FUNCTION "LGF_MatrixInverse" : Void
{ S7_Optimized_Access := 'TRUE' }
AUTHOR : Siemens_Digital_Industry
FAMILY : LGF
NAME : LGF_MatrixInverse
   VAR_OUTPUT
      error : Bool;
      status : Word;
   END_VAR

   VAR_IN_OUT
      matrix : Array[*, *] of LReal;
      matrixResult : Array[*, *] of LReal;
   END_VAR

   VAR_TEMP
      tempMatrix1LowerBoundRows : DInt;
      tempMatrix1LowerBoundColumns : DInt;
      tempMatrix1UpperBoundRows : DInt;
      tempMatrix1UpperBoundColumns : DInt;
      tempResultMatrixLowerBoundRows : DInt;
      tempResultMatrixLowerBoundColumns : DInt;
      tempResultMatrixUpperBoundRows : DInt;
      tempResultMatrixUpperBoundColumns : DInt;
      tempCounterRows : DInt;
      tempCounterColumns : DInt;
      tempColumns : DInt;
      tempRows : DInt;
      tempK : DInt;
      tempI : DInt;
      tempJ : DInt;
      tempMatrixElement : LReal;
   END_VAR

   VAR CONSTANT
      PRECISION : LReal := 1.0E-10;
      NEGATIVE_NUMERATOR : LReal := -1.0;
      ZERO : UInt := 0;
      ONE : UInt := 1;
      ROWS : UInt := 1;
      COLUMNS : UInt := 2;
      STATUS_NO_ERROR : Word := 16#0000;
      ERR_NOT_SQUARE_MATRIX : Word := 16#8200;
      ERR_ALGORITHM_NOT_POSSIBLE : Word := 16#8201;
      ERR_MATR1_LOWBOUND_ROWS_RESMATR_LOWBOUND_ROWS : Word := 16#8202;
      ERR_MATR1_LOWBOUND_COLUMNS_RESMATR_LOWBOUND_COLUMNS : Word := 16#8203;
      ERR_MATR1_UPPBOUND_ROWS_RESMATR_UPPBOUND_ROWS : Word := 16#8204;
      ERR_MATR1_UPPBOUND_COLUMNS_RESMATR_UPPBOUND_COLUMNS : Word := 16#8205;
   END_VAR


BEGIN
	REGION Block info header
	  //=============================================================================
	  // SIEMENS AG / (c)Copyright 2017
	  //-------------------------------------------------------------------------------
	  // Title:            LGF_MatrixInverse
	  // Comment/Function: Caluclates an inverted version of a matrix
	  // Library/Family:   LGF(Library General Functions)
	  // Author:           Siemens Digital Industry Support
	  // Tested with:      S7-PLCSIM Advanced V2.0 SP1
	  // Engineering:      TIA Portal V15 Update 2
	  // Restrictions:     ENO disabled - error handling done by error and status
	  // Requirements:     PLC (S7-1200 / S7-1500)
	  //-------------------------------------------------------------------------------
	  //=================================================================================
	END_REGION Block info header

	REGION Determine the size of the matrices
	  // Lower bound rows
	  #tempMatrix1LowerBoundRows := LOWER_BOUND(ARR := #matrix, DIM := #ROWS);
	  #tempResultMatrixLowerBoundRows := LOWER_BOUND(ARR := #matrixResult, DIM := #ROWS);
	  // Lower bound columns
	  #tempMatrix1LowerBoundColumns := LOWER_BOUND(ARR := #matrix, DIM := #COLUMNS);
	  #tempResultMatrixLowerBoundColumns := LOWER_BOUND(ARR := #matrixResult, DIM := #COLUMNS);
	  // Upper bound rows
	  #tempMatrix1UpperBoundRows := UPPER_BOUND(ARR := #matrix, DIM := #ROWS);
	  #tempResultMatrixUpperBoundRows := UPPER_BOUND(ARR := #matrixResult, DIM := #ROWS);
	  // Upper bound columns
	  #tempMatrix1UpperBoundColumns := UPPER_BOUND(ARR := #matrix, DIM := #COLUMNS);
	  #tempResultMatrixUpperBoundColumns := UPPER_BOUND(ARR := #matrixResult, DIM := #COLUMNS);
	END_REGION

	REGION Count the columns and rows of input matrix
	  // Count the columns
	  IF #tempMatrix1LowerBoundColumns = #ZERO THEN
	    #tempColumns := #tempMatrix1UpperBoundColumns + #ONE;
	  ELSE
	    #tempColumns := (#tempMatrix1UpperBoundColumns - #tempMatrix1LowerBoundColumns) + #ONE;
	  END_IF;
	  // Count the rows
	  IF #tempMatrix1LowerBoundRows = #ZERO THEN
	    #tempRows := #tempMatrix1UpperBoundRows + #ONE;
	  ELSE
	    #tempRows := (#tempMatrix1UpperBoundRows - #tempMatrix1LowerBoundRows) + #ONE;
	  END_IF;
	END_REGION

	REGION Error validation
	  // Check whether input matrix is a square matrix
	  IF #tempRows <> #tempColumns THEN
	    #error := TRUE;
	    #status := #ERR_NOT_SQUARE_MATRIX;
	    RETURN;
	  END_IF;

	  // Output matrix must have same lower bounds as the input matrix. (Same array size)
	  IF (#tempMatrix1LowerBoundRows <> #tempResultMatrixLowerBoundRows) THEN
	    #error := TRUE;
	    #status := #ERR_MATR1_LOWBOUND_ROWS_RESMATR_LOWBOUND_ROWS;
	    RETURN;
	  ELSIF (#tempMatrix1LowerBoundColumns <> #tempResultMatrixLowerBoundColumns) THEN
	    #error := TRUE;
	    #status := #ERR_MATR1_LOWBOUND_COLUMNS_RESMATR_LOWBOUND_COLUMNS;
	    RETURN;
	  END_IF;
	  // Output matrix must have same upper bounds as the input matrix. (Same array size)
	  IF (#tempMatrix1UpperBoundRows <> #tempResultMatrixUpperBoundRows) THEN
	    #error := TRUE;
	    #status := #ERR_MATR1_UPPBOUND_ROWS_RESMATR_UPPBOUND_ROWS;
	    RETURN;
	  ELSIF (#tempMatrix1UpperBoundColumns <> #tempResultMatrixUpperBoundColumns) THEN
	    #error := TRUE;
	    #status := #ERR_MATR1_UPPBOUND_COLUMNS_RESMATR_UPPBOUND_COLUMNS;
	    RETURN;
	  END_IF;
	END_REGION

	REGION Calculation of the inversed matrix
	  #matrixResult[#tempMatrix1LowerBoundRows, #tempMatrix1LowerBoundColumns] := #ZERO;
	  // Negate the input matrix and copy to output matrix.
	  FOR #tempCounterRows := #tempMatrix1LowerBoundRows TO #tempMatrix1UpperBoundRows DO
	    FOR #tempCounterColumns := #tempMatrix1LowerBoundColumns TO #tempMatrix1UpperBoundColumns DO
	      #matrixResult[#tempCounterRows, #tempCounterColumns] := - #matrix[#tempCounterRows, #tempCounterColumns];
	    END_FOR;
	  END_FOR;

	  //Outside loop - relegation of "Main" diagonal
	  FOR #tempK := #tempMatrix1LowerBoundColumns TO #tempMatrix1UpperBoundColumns DO
	    // Avoid a division by zero --> Error: Algorithm does not work for the input matrix.

	    #tempMatrixElement := #matrixResult[#tempK, #tempK];
	    IF ABS(#tempMatrixElement - #ZERO) <= (#PRECISION * ABS(#tempMatrixElement)) THEN
	      #error := TRUE;
	      #status := #ERR_ALGORITHM_NOT_POSSIBLE;
	      RETURN;
	    END_IF;

	    //Calculation of Pivot-element
	    #tempMatrixElement := (#NEGATIVE_NUMERATOR / #tempMatrixElement);
	    #matrixResult[#tempK, #tempK] := #tempMatrixElement;

	    //Calculation of elemente in the Pivot-column.
	    FOR #tempI := #tempMatrix1LowerBoundColumns TO #tempMatrix1UpperBoundColumns DO
	      IF #tempI <> #tempK THEN
	        #matrixResult[#tempI, #tempK] :=
	        #matrixResult[#tempI, #tempK] * #matrixResult[#tempK, #tempK];
	      END_IF;
	    END_FOR;

	    // Convert-calculation of elements, which are NOT in the Pivot-rolumn AND NOT in the Pivot-row.
	    FOR #tempI := #tempMatrix1LowerBoundRows TO #tempMatrix1UpperBoundRows DO
	      IF #tempI <> #tempK THEN
	        FOR #tempJ := #tempMatrix1LowerBoundColumns TO #tempMatrix1UpperBoundColumns DO
	          IF #tempJ <> #tempK THEN
	            #matrixResult[#tempI, #tempJ] :=
	            #matrixResult[#tempI, #tempJ] + #matrixResult[#tempI, #tempK] * #matrixResult[#tempK, #tempJ];
	          END_IF;
	        END_FOR;
	      END_IF;
	    END_FOR;

	    //Calculation of elements in the Pivot-row.
	    FOR #tempJ := #tempMatrix1LowerBoundColumns TO #tempMatrix1UpperBoundColumns DO
	      IF #tempJ <> #tempK THEN
	        #matrixResult[#tempK, #tempJ] :=
	        #matrixResult[#tempK, #tempJ] * #matrixResult[#tempK, #tempK];
	      END_IF;
	    END_FOR;
	  END_FOR;

	  #error := false;
	  #status := #STATUS_NO_ERROR;
	  // ENO mechanism is not used
	  ENO := TRUE;
	END_REGION

END_FUNCTION